TEXTLIST TextList_Piston_Recipe_State_DownUp
  0 = ' '
  1 = 'Down'
  2 = 'Up'
   = ''
END_TEXTLIST

(* stored: Version 1.1.0.1, ProductVersion 3.1.4024.12
   TextList TextList_Piston_Recipe_State_DownUp: Id {871bc978-8184-418b-a96b-42bce59c1583} *)
